TYPE ST_PolarIIChamber_HolderServiceParam :
STRUCT
	Gripper : ST_PolarIIChamber_OpenCloseServiceParam;
	Rotate : ST_PolarIIChamber_HolderRotateServiceParam;
	VacuumEstablish : ST_EmptyServiceParam;
END_STRUCT
END_TYPE

(* stored: Version 1.1.0.1, ProductVersion 3.1.4026.18
   DUT ST_PolarIIChamber_HolderServiceParam: Id {14000000-0000-0000-0000-000000000065} *)
